Fanuc KAREL source: KT00290.KL

PROGRAM KT00290
%NOLOCKGROUP
VAR
  P1: JOINTPOS
  P2: JOINTPOS
  OUT: BOOLEAN
BEGIN
  OUT = P1 = P2
END KT00290
